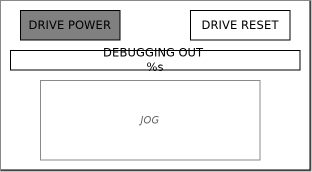
VISUALIZATION DRIVE  // 312x172
    Rectangle (0,0 310x170)
    Rectangle (10,50 290x20), "DEBUGGING OUT %s", text variable: MAIN.Track.eState
    Rectangle (20,10 100x30), "DRIVE POWER", colour toggle: MAIN.Track.Enable
    Rectangle (190,10 100x30), "DRIVE RESET", colour toggle: MAIN.Track.ResetBit
        tap MAIN.Track.ResetBit
    Frame (40,80 220x80)
        shows JOG()
END_VISUALIZATION

(* stored: Version 1.1.0.1, ProductVersion 3.1.4024.16
   Visu DRIVE: Id {7527a4bf-4007-4b0a-b018-21db365d173f} *)
